Staubli VAL3: new.pgx

public program new()
  local string l_sPage
  local bool l_bExit
  local num l_i
  local num l_nToolIndex
  local num l_nFrameIndex
  local bool l_bResult
  local bool l_bResult1
  local num l_nSize
  local string l_sHeader
  local num l_nID
  local bool l_bFound
begin
  // l_sPage=""
  do
    if util:sPage!="new"
      util:sPage="new"
      resize(sFrameList,1,size(saveData:fFrameItem))
      resize(sToolList,1,size(saveData:tToolItem))
      for l_i = 0 to size(sFrameList)-1
        sFrameList[l_i]=toString("",l_i)+","+saveData:fFrameItem[l_i].sName
      endFor
      for l_i = 0 to size(sToolList)-1
        sToolList[l_i]=toString("",l_i)+","+saveData:tToolItem[l_i].sName
      endFor
      sNewName=""
      nMoveID=0
      bCancel=false
      bConfirm=false
      sSelFrame=""
      sSelTool=""
      userPageBind("new","txt1","value",sNewName,1,"rw")
      userPageBind("new","nmb1","value",nMoveID,1,"rw")
      userPageBind("new","cbx1","options",sFrameList,size(sFrameList),"r")
      userPageBind("new","cbx2","options",sToolList,size(sToolList),"r")
      userPageBind("new","cbx1","value",sSelFrame,1,"rw")
      userPageBind("new","cbx2","value",sSelTool,1,"rw")
      userPageBindClick("new","btn1",bConfirm,true)
      userPageBindClick("new","btn2",bCancel,true)
      userPage(util:sPage)
      delay(0.5)

    endIf
    //
    toNum(sSelFrame,l_nFrameIndex,l_bResult)
    toNum(sSelTool,l_nToolIndex,l_bResult1)
    //button
    if bConfirm
      bConfirm=false
      if l_bResult and l_bResult1
        call trajectory:getSize(l_nSize)
        call getTrajID()
        l_nID=0
        do
          l_i=0
          do
            if l_nID==nIDIsExit[l_i]
              l_bFound=true
               l_nID=l_nID+1
            else
              l_bFound=false
            endIf
            l_i=l_i+1
          until l_bFound==false or l_i>=size(nIDIsExit)

          until l_bFound==false

        if l_nSize<10
          l_sHeader="0"+toString("",l_nID)+" "+sNewName
        else
          l_sHeader=toString("",l_nID)+" "+sNewName
        endIf
          call trajectory:new(l_sHeader,l_nFrameIndex,l_nToolIndex,nMoveID,bToSave)
          call trajectory:onSave(bToSave)
          sSelTraj=l_sHeader
          l_bExit=true
      else
        popUpMsg("设定的数据非法")
      endIf
    elseIf bCancel
      bCancel=false
      l_bExit=true
    endIf


    delay(0)
  until l_bExit==true

end
